(* IEC 61131-3 sources: llm-plc-st-eval/codesys/dobles/B5, 7 files *)

(* ---- 01_Correcta.st ---- *)
(* DOBLE DE PRUEBA B5/Correcta - NO ES CORPUS. Esperado: veredicto 1 *)
FUNCTION_BLOCK FB_Ventilador
VAR_INPUT
    quemadorOn : BOOL;
END_VAR
VAR_OUTPUT
    ventilador : BOOL;
END_VAR
VAR
    t : TOF;
END_VAR
t(IN := quemadorOn, PT := T#30S);
ventilador := t.Q;
END_FUNCTION_BLOCK

(* ---- 02_TiempoCorto.st ---- *)
(* DOBLE DE PRUEBA B5/TiempoCorto - NO ES CORPUS. Esperado: veredicto 2, falla en el paso 2 *)
FUNCTION_BLOCK FB_Ventilador
VAR_INPUT
    quemadorOn : BOOL;
END_VAR
VAR_OUTPUT
    ventilador : BOOL;
END_VAR
VAR
    t : TOF;
END_VAR
t(IN := quemadorOn, PT := T#10S);
ventilador := t.Q;
END_FUNCTION_BLOCK

(* ---- 03_TiempoLargo.st ---- *)
(* DOBLE DE PRUEBA B5/TiempoLargo - NO ES CORPUS. Esperado: veredicto 2, falla en el paso 3 *)
FUNCTION_BLOCK FB_Ventilador
VAR_INPUT
    quemadorOn : BOOL;
END_VAR
VAR_OUTPUT
    ventilador : BOOL;
END_VAR
VAR
    t : TOF;
END_VAR
t(IN := quemadorOn, PT := T#60S);
ventilador := t.Q;
END_FUNCTION_BLOCK

(* ---- 04_SinRetardo.st ---- *)
(* DOBLE DE PRUEBA B5/SinRetardo - NO ES CORPUS. Esperado: veredicto 2, falla en el paso 2 *)
FUNCTION_BLOCK FB_Ventilador
VAR_INPUT
    quemadorOn : BOOL;
END_VAR
VAR_OUTPUT
    ventilador : BOOL;
END_VAR
VAR
    nada : BOOL;
END_VAR
ventilador := quemadorOn;
END_FUNCTION_BLOCK

(* ---- 05_TonEnVezDeTof.st ---- *)
(* DOBLE DE PRUEBA B5/TonEnVezDeTof - NO ES CORPUS. Esperado: veredicto 2, falla en el paso 1 *)
FUNCTION_BLOCK FB_Ventilador
VAR_INPUT
    quemadorOn : BOOL;
END_VAR
VAR_OUTPUT
    ventilador : BOOL;
END_VAR
VAR
    t : TON;
END_VAR
t(IN := quemadorOn, PT := T#30S);
ventilador := t.Q;
END_FUNCTION_BLOCK

(* ---- 06_SinRearme.st ---- *)
(* DOBLE DE PRUEBA B5/SinRearme - NO ES CORPUS. Esperado: veredicto 2, falla en el paso 5 *)
FUNCTION_BLOCK FB_Ventilador
VAR_INPUT
    quemadorOn : BOOL;
END_VAR
VAR_OUTPUT
    ventilador : BOOL;
END_VAR
VAR
    tAhora : TIME;
    tPrev : TIME;
    dScan : TIME;
    init : BOOL;
    acum : TIME;
END_VAR
tAhora := TIME();
IF NOT init THEN
    tPrev := tAhora;
    init := TRUE;
END_IF
dScan := tAhora - tPrev;
tPrev := tAhora;
IF quemadorOn THEN
    ventilador := TRUE;          (* no reinicia el acumulador *)
ELSE
    acum := acum + dScan;
    IF acum >= T#30S THEN
        ventilador := FALSE;
    END_IF
END_IF
END_FUNCTION_BLOCK

(* ---- 07_RearmeCorto.st ---- *)
(* DOBLE DE PRUEBA B5/RearmeCorto - NO ES CORPUS. Esperado: veredicto 2, falla en el paso 7 *)
FUNCTION_BLOCK FB_Ventilador
VAR_INPUT
    quemadorOn : BOOL;
END_VAR
VAR_OUTPUT
    ventilador : BOOL;
END_VAR
VAR
    tAhora : TIME;
    tPrev : TIME;
    dScan : TIME;
    init : BOOL;
    acum : TIME;
    ciclos : INT;
    prev : BOOL;
    pt : TIME;
END_VAR
tAhora := TIME();
IF NOT init THEN
    tPrev := tAhora;
    init := TRUE;
END_IF
dScan := tAhora - tPrev;
tPrev := tAhora;
IF quemadorOn THEN
    ventilador := TRUE;
    acum := T#0S;
ELSE
    IF prev THEN
        ciclos := ciclos + 1;    (* flanco de bajada del quemador *)
    END_IF
    acum := acum + dScan;
    IF ciclos <= 1 THEN
        pt := T#30S;
    ELSE
        pt := T#15S;
    END_IF
    IF acum >= pt THEN
        ventilador := FALSE;
    END_IF
END_IF
prev := quemadorOn;
END_FUNCTION_BLOCK
